SUBAPPLICATION INI_IN_AND_STORE_AUDI2_OVERRIDE (* Wie INI_IN_AND_STORE_AUDI2, aber MIT Override-Moeglichkeit: Socket OVERRIDE_ACTIVE (AX) erzwingt bei TRUE kontinuierlich einen konfigurierten Wert (Default 1=Deaktiviert) statt des Live-VT-Werts - z.B. fuer gegenseitigen Options-Ausschluss. Bei OVERRIDE_ACTIVE=FALSE (unbenutzt) identisches Verhalten wie INI_IN_AND_STORE_AUDI2. *)
  (* Standard: 61499-2; Description: Copyright (c) 2026 Meisterschulen am Ostbahnhof This program and the accompanying materials are made available under the terms of the Eclipse Public License 2.0 which is available at https://www.eclipse.org/legal/epl-2.0/ SPDX-License-Identifier: EPL-2.0 *)
  (* Version 1.2, 2026-10-13, Franz Höpfinger, Meisterschulen am Ostbahnhof, Umbenannt von INI_IN_AND_STORE_AUDI2 zu INI_IN_AND_STORE_AUDI2_OVERRIDE, damit der Name die Override-Moeglichkeit klar erkennen laesst. Die schlanke Variante ohne OVERRIDE_ACTIVE-Socket (fuer Aufrufer, die ihn nicht brauchen) liegt jetzt separat unter INI_IN_AND_STORE_AUDI2. *)
  (* Version 1.1, 2026-10-13, Franz Höpfinger, Meisterschulen am Ostbahnhof, Neuer Socket OVERRIDE_ACTIVE (AX, Default unbenutzt/FALSE) - erzwingt bei TRUE kontinuierlich VAL=1 (Deaktiviert) statt des Live-VT-Werts, ueber SEL_Override (AUDI_AX_SEL_AUDI) vor AUDI_TO_AUDI2 eingefuegt. Laeuft ueber denselben bestehenden INI_AUDI2/Q_NumericValue_AUDI-Pfad - Q_NumericValue erlaubt laut eigener Doku nur eine Instanz je ObjId, daher keine zweite Schreib-Instanz moeglich. Fuer gegenseitigen Options-Ausschluss (BunkerKlappen/AufnahmeRechts), unveraendertes Verhalten wenn unbenutzt. *)
  (* Version 1.0, 2026-10-11, Franz Höpfinger, Meisterschulen am Ostbahnhof, AUDI2 adapter variant of INI_IN_AND_STORE_AUDI - NumericValue_IDA + AD_TO_AUDI + AUDI_TO_AUDI2 + INI_AUDI2 (bidirektionaler Adapter statt AUDI+Split-Paar), AUDI_TO_AUDI2.AUDI_OUT gesplittet auf Q_NumericValue_AUDI (VT-Anzeige) und VALUEO (weiterer Consumer). Fuer reine Enum/Ganzzahl-Werte (z.B. Optionsseite Dropdowns 0-3), keine Dezimalstellen. *)
  PACKAGE MyLib::sys;
  IMPORT isobus::UT::Q::const::IDs::ID_NULL;
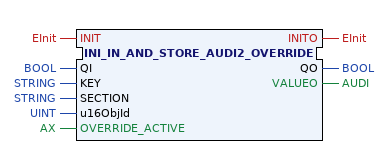
  EVENT_INPUT
    INIT : EInit; (* Initialization Request *)
  END_EVENT
  EVENT_OUTPUT
    INITO : EInit; (* Initialization Confirm *)
  END_EVENT
  VAR_INPUT
    QI : BOOL := TRUE; (* Quality Input - TRUE to enable service *)
    KEY : STRING; (* Key name. *)
    SECTION : STRING; (* Section name. *)
    u16ObjId : UINT := ID_NULL;
  END_VAR
  VAR_OUTPUT
    QO : BOOL; (* Quality Output - TRUE if service executed successfully *)
  END_VAR
  SOCKETS
    OVERRIDE_ACTIVE : adapter::types::unidirectional::AX; (* Kontinuierlich TRUE erzwingt VAL=1 (Deaktiviert), unabhaengig vom Live-VT-Wert - fuer gegenseitigen Options-Ausschluss. FALSE (unbenutzt, Default bei den meisten Aufrufern) = unveraendertes Verhalten. *)
  END_SOCKETS
  PLUGS
    VALUEO : adapter::types::unidirectional::AUDI;
  END_PLUGS
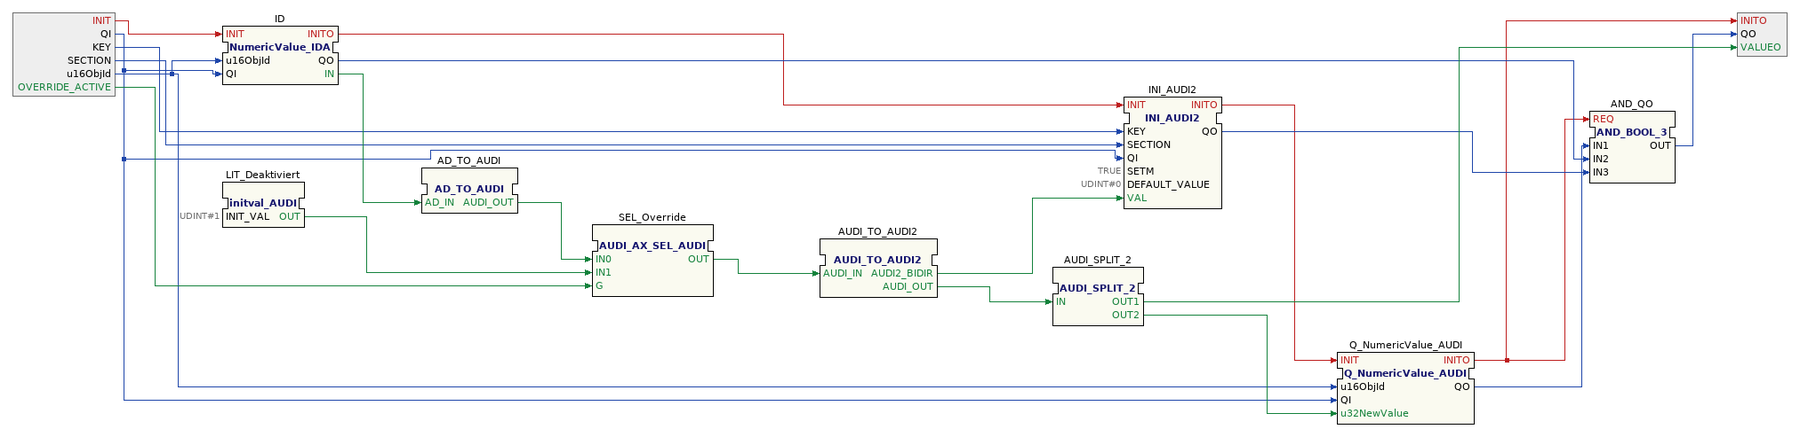
  (* SETM=TRUE - der Boot-Wert laedt so oder so automatisch (INIT -> INITO -> GET -> GETO, unabhaengig von SETM). SETM=TRUE sorgt dafuer, dass auch eine LIVE-Aenderung waehrend des laufenden Betriebs sofort bestaetigt/zurueckgemeldet wird - wichtig, falls der frische Wert noch im selben Lauf weiterverwendet werden soll (z.B. hier ueber VALUEO). *)
  FBS
    ID : isobus::UT::io::NumericValue::NumericValue_IDA;
    AD_TO_AUDI : adapter::conversion::unidirectional::AD_TO_AUDI;
    LIT_Deaktiviert : adapter::types::unidirectional::AUDI::initval::initval_AUDI(INIT_VAL := UDINT#1); (* Override-Wert: 1=Deaktiviert *)
    SEL_Override : adapter::iec61131::selection::AUDI_AX_SEL_AUDI; (* IN0=Live-VT-Wert (unveraendert), IN1=Deaktiviert-Override, G=OVERRIDE_ACTIVE *)
    AUDI_TO_AUDI2 : adapter::conversion::bidirectional::AUDI_TO_AUDI2;
    INI_AUDI2 : eclipse4diac::storage::INI_AUDI2(SETM := TRUE, DEFAULT_VALUE := UDINT#0);
    AUDI_SPLIT_2 : adapter::events::unidirectional::AUDI_SPLIT_2;
    Q_NumericValue_AUDI : isobus::UT::Q::Q_NumericValue_AUDI;
    AND_QO : iec61131::booleanOperators::AND_BOOL_3;
  END_FBS
  EVENT_CONNECTIONS
    INIT TO ID.INIT;
    ID.INITO TO INI_AUDI2.INIT;
    INI_AUDI2.INITO TO Q_NumericValue_AUDI.INIT;
    Q_NumericValue_AUDI.INITO TO INITO;
    Q_NumericValue_AUDI.INITO TO AND_QO.REQ;
  END_CONNECTIONS
  DATA_CONNECTIONS
    KEY TO INI_AUDI2.KEY;
    SECTION TO INI_AUDI2.SECTION;
    u16ObjId TO ID.u16ObjId;
    u16ObjId TO Q_NumericValue_AUDI.u16ObjId;
    QI TO Q_NumericValue_AUDI.QI;
    QI TO ID.QI;
    QI TO INI_AUDI2.QI;
    Q_NumericValue_AUDI.QO TO AND_QO.IN1;
    ID.QO TO AND_QO.IN2;
    INI_AUDI2.QO TO AND_QO.IN3;
    AND_QO.OUT TO QO;
  END_CONNECTIONS
  ADAPTER_CONNECTIONS
    ID.IN TO AD_TO_AUDI.AD_IN;
    AD_TO_AUDI.AUDI_OUT TO SEL_Override.IN0;
    LIT_Deaktiviert.OUT TO SEL_Override.IN1;
    OVERRIDE_ACTIVE TO SEL_Override.G;
    SEL_Override.OUT TO AUDI_TO_AUDI2.AUDI_IN;
    AUDI_TO_AUDI2.AUDI2_BIDIR TO INI_AUDI2.VAL;
    AUDI_TO_AUDI2.AUDI_OUT TO AUDI_SPLIT_2.IN;
    AUDI_SPLIT_2.OUT1 TO VALUEO;
    AUDI_SPLIT_2.OUT2 TO Q_NumericValue_AUDI.u32NewValue;
  END_CONNECTIONS
END_SUBAPPLICATION
